Staubli VAL3: CalAdjustXY2.pgx

public program CalAdjustXY2()
  local trsf l_trFlange
  local trsf l_trTCP
  local num x
  local num y
  local num z
begin
  //初始化数据
  l_trFlange={0,0,0,0,0,0}
  l_trTCP={0,0,0,0,0,0}
  //计算新的中心位置
  x=(db:pAdjustXY_2_1.trsf.x+db:pAdjustXY_2_2.trsf.x)/2
  y=(db:pAdjustXY_2_1.trsf.y+db:pAdjustXY_2_2.trsf.y)/2
  z=db:pAdjustXY_2_1.trsf.z
  //
  l_trFlange=db:pAdjustXY_2_1.trsf*!db:utCurrentTool.tValue.trsf
  if db:sMounting=="Floor"
    l_trTCP={x,y,z,0,180,0}
  elseIf db:sMounting=="Ceiling"
    l_trTCP={x,y,z,0,0,0}
  endIf
  db:tTool2.trsf=!l_trFlange*l_trTCP
  //
  db:tTool2.trsf.rx=db:tTool1.trsf.rx
  db:tTool2.trsf.ry=db:tTool1.trsf.ry
  db:tTool2.trsf.rz=db:tTool1.trsf.rz
  call db:hmiAlert("SaveInTool2","info")
end
